Fanuc KAREL source: KA00076.KL

PROGRAM KA00076
%NOLOCKGROUP
VAR
  SRC: XYZWPREXT
  DST: STRING[80]
BEGIN
  SRC.X = 1.0
  DST = SRC
END KA00076
